// TIA Portal V19 export
DATA_BLOCK "ALL HOOTER_DB"   // DB1
// stored: InstanceOfName ALL HOOTER, InstanceOfType FB
"ALL HOOTER"
   // VAR
   //    HOOTER_Instance { S7_SetPoint := 'True'} : "HOOTER";
   //    HOOTER_Instance_1 { S7_SetPoint := 'True'} : "HOOTER";
   // END_VAR
BEGIN
END_DATA_BLOCK
